(* IEC 61131-3 sources: STAR-PLC-Agent/results/raw/codex_matrix_resume_20261114/codex_deepseek/SELF010/functional/attempt_0001, 1 file *)

(* ---- test_program.st ---- *)
PROGRAM PLC_PRG
VAR
 BenchStep : UDINT := 0;
 BenchCalls : UDINT := 0;
 BenchDone : BOOL := FALSE;
 BenchUut0 : FB_Task;
 BenchUut1 : FB_Task;
 BenchUut2 : FB_Task;
 BenchUut3 : FB_Task;
 BenchUut4 : FB_Task;
 BenchUut5 : FB_Task;
 BenchUut6 : FB_Task;
 BenchUut7 : FB_Task;
 TraceIn_Fault : ARRAY[0..49] OF BOOL;
 TraceIn_Ack : ARRAY[0..49] OF BOOL;
 TraceIn_Reset : ARRAY[0..49] OF BOOL;
 TraceOut_Alarm : ARRAY[0..49] OF BOOL;
 TraceOut_Acknowledged : ARRAY[0..49] OF BOOL;
 TraceOut_Horn : ARRAY[0..49] OF BOOL;
END_VAR

IF NOT BenchDone THEN
 CASE BenchStep OF
 0:
   BenchUut0.Fault := FALSE;
   BenchUut0.Ack := FALSE;
   BenchUut0.Reset := FALSE;
   TraceIn_Fault[0] := BenchUut0.Fault;
   TraceIn_Ack[0] := BenchUut0.Ack;
   TraceIn_Reset[0] := BenchUut0.Reset;
   BenchUut0();
   TraceOut_Alarm[0] := BenchUut0.Alarm;
   TraceOut_Acknowledged[0] := BenchUut0.Acknowledged;
   TraceOut_Horn[0] := BenchUut0.Horn;
   BenchCalls := BenchCalls + 1;
 1:
   BenchUut0.Fault := TRUE;
   BenchUut0.Ack := TRUE;
   BenchUut0.Reset := FALSE;
   TraceIn_Fault[1] := BenchUut0.Fault;
   TraceIn_Ack[1] := BenchUut0.Ack;
   TraceIn_Reset[1] := BenchUut0.Reset;
   BenchUut0();
   TraceOut_Alarm[1] := BenchUut0.Alarm;
   TraceOut_Acknowledged[1] := BenchUut0.Acknowledged;
   TraceOut_Horn[1] := BenchUut0.Horn;
   BenchCalls := BenchCalls + 1;
 2:
   BenchUut0.Fault := TRUE;
   BenchUut0.Ack := TRUE;
   BenchUut0.Reset := FALSE;
   TraceIn_Fault[2] := BenchUut0.Fault;
   TraceIn_Ack[2] := BenchUut0.Ack;
   TraceIn_Reset[2] := BenchUut0.Reset;
   BenchUut0();
   TraceOut_Alarm[2] := BenchUut0.Alarm;
   TraceOut_Acknowledged[2] := BenchUut0.Acknowledged;
   TraceOut_Horn[2] := BenchUut0.Horn;
   BenchCalls := BenchCalls + 1;
 3:
   BenchUut0.Fault := FALSE;
   BenchUut0.Ack := FALSE;
   BenchUut0.Reset := FALSE;
   TraceIn_Fault[3] := BenchUut0.Fault;
   TraceIn_Ack[3] := BenchUut0.Ack;
   TraceIn_Reset[3] := BenchUut0.Reset;
   BenchUut0();
   TraceOut_Alarm[3] := BenchUut0.Alarm;
   TraceOut_Acknowledged[3] := BenchUut0.Acknowledged;
   TraceOut_Horn[3] := BenchUut0.Horn;
   BenchCalls := BenchCalls + 1;
 4:
   BenchUut0.Fault := TRUE;
   BenchUut0.Ack := FALSE;
   BenchUut0.Reset := FALSE;
   TraceIn_Fault[4] := BenchUut0.Fault;
   TraceIn_Ack[4] := BenchUut0.Ack;
   TraceIn_Reset[4] := BenchUut0.Reset;
   BenchUut0();
   TraceOut_Alarm[4] := BenchUut0.Alarm;
   TraceOut_Acknowledged[4] := BenchUut0.Acknowledged;
   TraceOut_Horn[4] := BenchUut0.Horn;
   BenchCalls := BenchCalls + 1;
 5:
   BenchUut0.Fault := FALSE;
   BenchUut0.Ack := FALSE;
   BenchUut0.Reset := TRUE;
   TraceIn_Fault[5] := BenchUut0.Fault;
   TraceIn_Ack[5] := BenchUut0.Ack;
   TraceIn_Reset[5] := BenchUut0.Reset;
   BenchUut0();
   TraceOut_Alarm[5] := BenchUut0.Alarm;
   TraceOut_Acknowledged[5] := BenchUut0.Acknowledged;
   TraceOut_Horn[5] := BenchUut0.Horn;
   BenchCalls := BenchCalls + 1;
 6:
   BenchUut1.Fault := TRUE;
   BenchUut1.Ack := FALSE;
   BenchUut1.Reset := TRUE;
   TraceIn_Fault[6] := BenchUut1.Fault;
   TraceIn_Ack[6] := BenchUut1.Ack;
   TraceIn_Reset[6] := BenchUut1.Reset;
   BenchUut1();
   TraceOut_Alarm[6] := BenchUut1.Alarm;
   TraceOut_Acknowledged[6] := BenchUut1.Acknowledged;
   TraceOut_Horn[6] := BenchUut1.Horn;
   BenchCalls := BenchCalls + 1;
 7:
   BenchUut1.Fault := TRUE;
   BenchUut1.Ack := TRUE;
   BenchUut1.Reset := TRUE;
   TraceIn_Fault[7] := BenchUut1.Fault;
   TraceIn_Ack[7] := BenchUut1.Ack;
   TraceIn_Reset[7] := BenchUut1.Reset;
   BenchUut1();
   TraceOut_Alarm[7] := BenchUut1.Alarm;
   TraceOut_Acknowledged[7] := BenchUut1.Acknowledged;
   TraceOut_Horn[7] := BenchUut1.Horn;
   BenchCalls := BenchCalls + 1;
 8:
   BenchUut1.Fault := FALSE;
   BenchUut1.Ack := TRUE;
   BenchUut1.Reset := TRUE;
   TraceIn_Fault[8] := BenchUut1.Fault;
   TraceIn_Ack[8] := BenchUut1.Ack;
   TraceIn_Reset[8] := BenchUut1.Reset;
   BenchUut1();
   TraceOut_Alarm[8] := BenchUut1.Alarm;
   TraceOut_Acknowledged[8] := BenchUut1.Acknowledged;
   TraceOut_Horn[8] := BenchUut1.Horn;
   BenchCalls := BenchCalls + 1;
 9:
   BenchUut2.Fault := TRUE;
   BenchUut2.Ack := FALSE;
   BenchUut2.Reset := TRUE;
   TraceIn_Fault[9] := BenchUut2.Fault;
   TraceIn_Ack[9] := BenchUut2.Ack;
   TraceIn_Reset[9] := BenchUut2.Reset;
   BenchUut2();
   TraceOut_Alarm[9] := BenchUut2.Alarm;
   TraceOut_Acknowledged[9] := BenchUut2.Acknowledged;
   TraceOut_Horn[9] := BenchUut2.Horn;
   BenchCalls := BenchCalls + 1;
 10:
   BenchUut2.Fault := TRUE;
   BenchUut2.Ack := TRUE;
   BenchUut2.Reset := TRUE;
   TraceIn_Fault[10] := BenchUut2.Fault;
   TraceIn_Ack[10] := BenchUut2.Ack;
   TraceIn_Reset[10] := BenchUut2.Reset;
   BenchUut2();
   TraceOut_Alarm[10] := BenchUut2.Alarm;
   TraceOut_Acknowledged[10] := BenchUut2.Acknowledged;
   TraceOut_Horn[10] := BenchUut2.Horn;
   BenchCalls := BenchCalls + 1;
 11:
   BenchUut2.Fault := TRUE;
   BenchUut2.Ack := TRUE;
   BenchUut2.Reset := TRUE;
   TraceIn_Fault[11] := BenchUut2.Fault;
   TraceIn_Ack[11] := BenchUut2.Ack;
   TraceIn_Reset[11] := BenchUut2.Reset;
   BenchUut2();
   TraceOut_Alarm[11] := BenchUut2.Alarm;
   TraceOut_Acknowledged[11] := BenchUut2.Acknowledged;
   TraceOut_Horn[11] := BenchUut2.Horn;
   BenchCalls := BenchCalls + 1;
 12:
   BenchUut3.Fault := FALSE;
   BenchUut3.Ack := TRUE;
   BenchUut3.Reset := FALSE;
   TraceIn_Fault[12] := BenchUut3.Fault;
   TraceIn_Ack[12] := BenchUut3.Ack;
   TraceIn_Reset[12] := BenchUut3.Reset;
   BenchUut3();
   TraceOut_Alarm[12] := BenchUut3.Alarm;
   TraceOut_Acknowledged[12] := BenchUut3.Acknowledged;
   TraceOut_Horn[12] := BenchUut3.Horn;
   BenchCalls := BenchCalls + 1;
 13:
   BenchUut3.Fault := TRUE;
   BenchUut3.Ack := FALSE;
   BenchUut3.Reset := FALSE;
   TraceIn_Fault[13] := BenchUut3.Fault;
   TraceIn_Ack[13] := BenchUut3.Ack;
   TraceIn_Reset[13] := BenchUut3.Reset;
   BenchUut3();
   TraceOut_Alarm[13] := BenchUut3.Alarm;
   TraceOut_Acknowledged[13] := BenchUut3.Acknowledged;
   TraceOut_Horn[13] := BenchUut3.Horn;
   BenchCalls := BenchCalls + 1;
 14:
   BenchUut3.Fault := FALSE;
   BenchUut3.Ack := FALSE;
   BenchUut3.Reset := FALSE;
   TraceIn_Fault[14] := BenchUut3.Fault;
   TraceIn_Ack[14] := BenchUut3.Ack;
   TraceIn_Reset[14] := BenchUut3.Reset;
   BenchUut3();
   TraceOut_Alarm[14] := BenchUut3.Alarm;
   TraceOut_Acknowledged[14] := BenchUut3.Acknowledged;
   TraceOut_Horn[14] := BenchUut3.Horn;
   BenchCalls := BenchCalls + 1;
 15:
   BenchUut3.Fault := FALSE;
   BenchUut3.Ack := TRUE;
   BenchUut3.Reset := FALSE;
   TraceIn_Fault[15] := BenchUut3.Fault;
   TraceIn_Ack[15] := BenchUut3.Ack;
   TraceIn_Reset[15] := BenchUut3.Reset;
   BenchUut3();
   TraceOut_Alarm[15] := BenchUut3.Alarm;
   TraceOut_Acknowledged[15] := BenchUut3.Acknowledged;
   TraceOut_Horn[15] := BenchUut3.Horn;
   BenchCalls := BenchCalls + 1;
 16:
   BenchUut3.Fault := TRUE;
   BenchUut3.Ack := TRUE;
   BenchUut3.Reset := FALSE;
   TraceIn_Fault[16] := BenchUut3.Fault;
   TraceIn_Ack[16] := BenchUut3.Ack;
   TraceIn_Reset[16] := BenchUut3.Reset;
   BenchUut3();
   TraceOut_Alarm[16] := BenchUut3.Alarm;
   TraceOut_Acknowledged[16] := BenchUut3.Acknowledged;
   TraceOut_Horn[16] := BenchUut3.Horn;
   BenchCalls := BenchCalls + 1;
 17:
   BenchUut3.Fault := TRUE;
   BenchUut3.Ack := FALSE;
   BenchUut3.Reset := TRUE;
   TraceIn_Fault[17] := BenchUut3.Fault;
   TraceIn_Ack[17] := BenchUut3.Ack;
   TraceIn_Reset[17] := BenchUut3.Reset;
   BenchUut3();
   TraceOut_Alarm[17] := BenchUut3.Alarm;
   TraceOut_Acknowledged[17] := BenchUut3.Acknowledged;
   TraceOut_Horn[17] := BenchUut3.Horn;
   BenchCalls := BenchCalls + 1;
 18:
   BenchUut3.Fault := FALSE;
   BenchUut3.Ack := FALSE;
   BenchUut3.Reset := TRUE;
   TraceIn_Fault[18] := BenchUut3.Fault;
   TraceIn_Ack[18] := BenchUut3.Ack;
   TraceIn_Reset[18] := BenchUut3.Reset;
   BenchUut3();
   TraceOut_Alarm[18] := BenchUut3.Alarm;
   TraceOut_Acknowledged[18] := BenchUut3.Acknowledged;
   TraceOut_Horn[18] := BenchUut3.Horn;
   BenchCalls := BenchCalls + 1;
 19:
   BenchUut4.Fault := TRUE;
   BenchUut4.Ack := FALSE;
   BenchUut4.Reset := FALSE;
   TraceIn_Fault[19] := BenchUut4.Fault;
   TraceIn_Ack[19] := BenchUut4.Ack;
   TraceIn_Reset[19] := BenchUut4.Reset;
   BenchUut4();
   TraceOut_Alarm[19] := BenchUut4.Alarm;
   TraceOut_Acknowledged[19] := BenchUut4.Acknowledged;
   TraceOut_Horn[19] := BenchUut4.Horn;
   BenchCalls := BenchCalls + 1;
 20:
   BenchUut4.Fault := FALSE;
   BenchUut4.Ack := FALSE;
   BenchUut4.Reset := FALSE;
   TraceIn_Fault[20] := BenchUut4.Fault;
   TraceIn_Ack[20] := BenchUut4.Ack;
   TraceIn_Reset[20] := BenchUut4.Reset;
   BenchUut4();
   TraceOut_Alarm[20] := BenchUut4.Alarm;
   TraceOut_Acknowledged[20] := BenchUut4.Acknowledged;
   TraceOut_Horn[20] := BenchUut4.Horn;
   BenchCalls := BenchCalls + 1;
 21:
   BenchUut4.Fault := FALSE;
   BenchUut4.Ack := TRUE;
   BenchUut4.Reset := FALSE;
   TraceIn_Fault[21] := BenchUut4.Fault;
   TraceIn_Ack[21] := BenchUut4.Ack;
   TraceIn_Reset[21] := BenchUut4.Reset;
   BenchUut4();
   TraceOut_Alarm[21] := BenchUut4.Alarm;
   TraceOut_Acknowledged[21] := BenchUut4.Acknowledged;
   TraceOut_Horn[21] := BenchUut4.Horn;
   BenchCalls := BenchCalls + 1;
 22:
   BenchUut4.Fault := FALSE;
   BenchUut4.Ack := FALSE;
   BenchUut4.Reset := FALSE;
   TraceIn_Fault[22] := BenchUut4.Fault;
   TraceIn_Ack[22] := BenchUut4.Ack;
   TraceIn_Reset[22] := BenchUut4.Reset;
   BenchUut4();
   TraceOut_Alarm[22] := BenchUut4.Alarm;
   TraceOut_Acknowledged[22] := BenchUut4.Acknowledged;
   TraceOut_Horn[22] := BenchUut4.Horn;
   BenchCalls := BenchCalls + 1;
 23:
   BenchUut4.Fault := FALSE;
   BenchUut4.Ack := FALSE;
   BenchUut4.Reset := TRUE;
   TraceIn_Fault[23] := BenchUut4.Fault;
   TraceIn_Ack[23] := BenchUut4.Ack;
   TraceIn_Reset[23] := BenchUut4.Reset;
   BenchUut4();
   TraceOut_Alarm[23] := BenchUut4.Alarm;
   TraceOut_Acknowledged[23] := BenchUut4.Acknowledged;
   TraceOut_Horn[23] := BenchUut4.Horn;
   BenchCalls := BenchCalls + 1;
 24:
   BenchUut4.Fault := FALSE;
   BenchUut4.Ack := FALSE;
   BenchUut4.Reset := FALSE;
   TraceIn_Fault[24] := BenchUut4.Fault;
   TraceIn_Ack[24] := BenchUut4.Ack;
   TraceIn_Reset[24] := BenchUut4.Reset;
   BenchUut4();
   TraceOut_Alarm[24] := BenchUut4.Alarm;
   TraceOut_Acknowledged[24] := BenchUut4.Acknowledged;
   TraceOut_Horn[24] := BenchUut4.Horn;
   BenchCalls := BenchCalls + 1;
 25:
   BenchUut4.Fault := FALSE;
   BenchUut4.Ack := TRUE;
   BenchUut4.Reset := FALSE;
   TraceIn_Fault[25] := BenchUut4.Fault;
   TraceIn_Ack[25] := BenchUut4.Ack;
   TraceIn_Reset[25] := BenchUut4.Reset;
   BenchUut4();
   TraceOut_Alarm[25] := BenchUut4.Alarm;
   TraceOut_Acknowledged[25] := BenchUut4.Acknowledged;
   TraceOut_Horn[25] := BenchUut4.Horn;
   BenchCalls := BenchCalls + 1;
 26:
   BenchUut5.Fault := FALSE;
   BenchUut5.Ack := FALSE;
   BenchUut5.Reset := FALSE;
   TraceIn_Fault[26] := BenchUut5.Fault;
   TraceIn_Ack[26] := BenchUut5.Ack;
   TraceIn_Reset[26] := BenchUut5.Reset;
   BenchUut5();
   TraceOut_Alarm[26] := BenchUut5.Alarm;
   TraceOut_Acknowledged[26] := BenchUut5.Acknowledged;
   TraceOut_Horn[26] := BenchUut5.Horn;
   BenchCalls := BenchCalls + 1;
 27:
   BenchUut5.Fault := TRUE;
   BenchUut5.Ack := TRUE;
   BenchUut5.Reset := FALSE;
   TraceIn_Fault[27] := BenchUut5.Fault;
   TraceIn_Ack[27] := BenchUut5.Ack;
   TraceIn_Reset[27] := BenchUut5.Reset;
   BenchUut5();
   TraceOut_Alarm[27] := BenchUut5.Alarm;
   TraceOut_Acknowledged[27] := BenchUut5.Acknowledged;
   TraceOut_Horn[27] := BenchUut5.Horn;
   BenchCalls := BenchCalls + 1;
 28:
   BenchUut5.Fault := TRUE;
   BenchUut5.Ack := TRUE;
   BenchUut5.Reset := FALSE;
   TraceIn_Fault[28] := BenchUut5.Fault;
   TraceIn_Ack[28] := BenchUut5.Ack;
   TraceIn_Reset[28] := BenchUut5.Reset;
   BenchUut5();
   TraceOut_Alarm[28] := BenchUut5.Alarm;
   TraceOut_Acknowledged[28] := BenchUut5.Acknowledged;
   TraceOut_Horn[28] := BenchUut5.Horn;
   BenchCalls := BenchCalls + 1;
 29:
   BenchUut5.Fault := FALSE;
   BenchUut5.Ack := FALSE;
   BenchUut5.Reset := FALSE;
   TraceIn_Fault[29] := BenchUut5.Fault;
   TraceIn_Ack[29] := BenchUut5.Ack;
   TraceIn_Reset[29] := BenchUut5.Reset;
   BenchUut5();
   TraceOut_Alarm[29] := BenchUut5.Alarm;
   TraceOut_Acknowledged[29] := BenchUut5.Acknowledged;
   TraceOut_Horn[29] := BenchUut5.Horn;
   BenchCalls := BenchCalls + 1;
 30:
   BenchUut5.Fault := TRUE;
   BenchUut5.Ack := FALSE;
   BenchUut5.Reset := FALSE;
   TraceIn_Fault[30] := BenchUut5.Fault;
   TraceIn_Ack[30] := BenchUut5.Ack;
   TraceIn_Reset[30] := BenchUut5.Reset;
   BenchUut5();
   TraceOut_Alarm[30] := BenchUut5.Alarm;
   TraceOut_Acknowledged[30] := BenchUut5.Acknowledged;
   TraceOut_Horn[30] := BenchUut5.Horn;
   BenchCalls := BenchCalls + 1;
 31:
   BenchUut5.Fault := FALSE;
   BenchUut5.Ack := FALSE;
   BenchUut5.Reset := TRUE;
   TraceIn_Fault[31] := BenchUut5.Fault;
   TraceIn_Ack[31] := BenchUut5.Ack;
   TraceIn_Reset[31] := BenchUut5.Reset;
   BenchUut5();
   TraceOut_Alarm[31] := BenchUut5.Alarm;
   TraceOut_Acknowledged[31] := BenchUut5.Acknowledged;
   TraceOut_Horn[31] := BenchUut5.Horn;
   BenchCalls := BenchCalls + 1;
 32:
   BenchUut5.Fault := TRUE;
   BenchUut5.Ack := FALSE;
   BenchUut5.Reset := TRUE;
   TraceIn_Fault[32] := BenchUut5.Fault;
   TraceIn_Ack[32] := BenchUut5.Ack;
   TraceIn_Reset[32] := BenchUut5.Reset;
   BenchUut5();
   TraceOut_Alarm[32] := BenchUut5.Alarm;
   TraceOut_Acknowledged[32] := BenchUut5.Acknowledged;
   TraceOut_Horn[32] := BenchUut5.Horn;
   BenchCalls := BenchCalls + 1;
 33:
   BenchUut5.Fault := TRUE;
   BenchUut5.Ack := FALSE;
   BenchUut5.Reset := TRUE;
   TraceIn_Fault[33] := BenchUut5.Fault;
   TraceIn_Ack[33] := BenchUut5.Ack;
   TraceIn_Reset[33] := BenchUut5.Reset;
   BenchUut5();
   TraceOut_Alarm[33] := BenchUut5.Alarm;
   TraceOut_Acknowledged[33] := BenchUut5.Acknowledged;
   TraceOut_Horn[33] := BenchUut5.Horn;
   BenchCalls := BenchCalls + 1;
 34:
   BenchUut6.Fault := FALSE;
   BenchUut6.Ack := FALSE;
   BenchUut6.Reset := FALSE;
   TraceIn_Fault[34] := BenchUut6.Fault;
   TraceIn_Ack[34] := BenchUut6.Ack;
   TraceIn_Reset[34] := BenchUut6.Reset;
   BenchUut6();
   TraceOut_Alarm[34] := BenchUut6.Alarm;
   TraceOut_Acknowledged[34] := BenchUut6.Acknowledged;
   TraceOut_Horn[34] := BenchUut6.Horn;
   BenchCalls := BenchCalls + 1;
 35:
   BenchUut6.Fault := TRUE;
   BenchUut6.Ack := TRUE;
   BenchUut6.Reset := FALSE;
   TraceIn_Fault[35] := BenchUut6.Fault;
   TraceIn_Ack[35] := BenchUut6.Ack;
   TraceIn_Reset[35] := BenchUut6.Reset;
   BenchUut6();
   TraceOut_Alarm[35] := BenchUut6.Alarm;
   TraceOut_Acknowledged[35] := BenchUut6.Acknowledged;
   TraceOut_Horn[35] := BenchUut6.Horn;
   BenchCalls := BenchCalls + 1;
 36:
   BenchUut6.Fault := TRUE;
   BenchUut6.Ack := TRUE;
   BenchUut6.Reset := FALSE;
   TraceIn_Fault[36] := BenchUut6.Fault;
   TraceIn_Ack[36] := BenchUut6.Ack;
   TraceIn_Reset[36] := BenchUut6.Reset;
   BenchUut6();
   TraceOut_Alarm[36] := BenchUut6.Alarm;
   TraceOut_Acknowledged[36] := BenchUut6.Acknowledged;
   TraceOut_Horn[36] := BenchUut6.Horn;
   BenchCalls := BenchCalls + 1;
 37:
   BenchUut6.Fault := FALSE;
   BenchUut6.Ack := FALSE;
   BenchUut6.Reset := FALSE;
   TraceIn_Fault[37] := BenchUut6.Fault;
   TraceIn_Ack[37] := BenchUut6.Ack;
   TraceIn_Reset[37] := BenchUut6.Reset;
   BenchUut6();
   TraceOut_Alarm[37] := BenchUut6.Alarm;
   TraceOut_Acknowledged[37] := BenchUut6.Acknowledged;
   TraceOut_Horn[37] := BenchUut6.Horn;
   BenchCalls := BenchCalls + 1;
 38:
   BenchUut6.Fault := TRUE;
   BenchUut6.Ack := FALSE;
   BenchUut6.Reset := FALSE;
   TraceIn_Fault[38] := BenchUut6.Fault;
   TraceIn_Ack[38] := BenchUut6.Ack;
   TraceIn_Reset[38] := BenchUut6.Reset;
   BenchUut6();
   TraceOut_Alarm[38] := BenchUut6.Alarm;
   TraceOut_Acknowledged[38] := BenchUut6.Acknowledged;
   TraceOut_Horn[38] := BenchUut6.Horn;
   BenchCalls := BenchCalls + 1;
 39:
   BenchUut6.Fault := FALSE;
   BenchUut6.Ack := FALSE;
   BenchUut6.Reset := TRUE;
   TraceIn_Fault[39] := BenchUut6.Fault;
   TraceIn_Ack[39] := BenchUut6.Ack;
   TraceIn_Reset[39] := BenchUut6.Reset;
   BenchUut6();
   TraceOut_Alarm[39] := BenchUut6.Alarm;
   TraceOut_Acknowledged[39] := BenchUut6.Acknowledged;
   TraceOut_Horn[39] := BenchUut6.Horn;
   BenchCalls := BenchCalls + 1;
 40:
   BenchUut6.Fault := FALSE;
   BenchUut6.Ack := TRUE;
   BenchUut6.Reset := TRUE;
   TraceIn_Fault[40] := BenchUut6.Fault;
   TraceIn_Ack[40] := BenchUut6.Ack;
   TraceIn_Reset[40] := BenchUut6.Reset;
   BenchUut6();
   TraceOut_Alarm[40] := BenchUut6.Alarm;
   TraceOut_Acknowledged[40] := BenchUut6.Acknowledged;
   TraceOut_Horn[40] := BenchUut6.Horn;
   BenchCalls := BenchCalls + 1;
 41:
   BenchUut6.Fault := FALSE;
   BenchUut6.Ack := TRUE;
   BenchUut6.Reset := TRUE;
   TraceIn_Fault[41] := BenchUut6.Fault;
   TraceIn_Ack[41] := BenchUut6.Ack;
   TraceIn_Reset[41] := BenchUut6.Reset;
   BenchUut6();
   TraceOut_Alarm[41] := BenchUut6.Alarm;
   TraceOut_Acknowledged[41] := BenchUut6.Acknowledged;
   TraceOut_Horn[41] := BenchUut6.Horn;
   BenchCalls := BenchCalls + 1;
 42:
   BenchUut7.Fault := FALSE;
   BenchUut7.Ack := FALSE;
   BenchUut7.Reset := FALSE;
   TraceIn_Fault[42] := BenchUut7.Fault;
   TraceIn_Ack[42] := BenchUut7.Ack;
   TraceIn_Reset[42] := BenchUut7.Reset;
   BenchUut7();
   TraceOut_Alarm[42] := BenchUut7.Alarm;
   TraceOut_Acknowledged[42] := BenchUut7.Acknowledged;
   TraceOut_Horn[42] := BenchUut7.Horn;
   BenchCalls := BenchCalls + 1;
 43:
   BenchUut7.Fault := TRUE;
   BenchUut7.Ack := TRUE;
   BenchUut7.Reset := FALSE;
   TraceIn_Fault[43] := BenchUut7.Fault;
   TraceIn_Ack[43] := BenchUut7.Ack;
   TraceIn_Reset[43] := BenchUut7.Reset;
   BenchUut7();
   TraceOut_Alarm[43] := BenchUut7.Alarm;
   TraceOut_Acknowledged[43] := BenchUut7.Acknowledged;
   TraceOut_Horn[43] := BenchUut7.Horn;
   BenchCalls := BenchCalls + 1;
 44:
   BenchUut7.Fault := TRUE;
   BenchUut7.Ack := TRUE;
   BenchUut7.Reset := FALSE;
   TraceIn_Fault[44] := BenchUut7.Fault;
   TraceIn_Ack[44] := BenchUut7.Ack;
   TraceIn_Reset[44] := BenchUut7.Reset;
   BenchUut7();
   TraceOut_Alarm[44] := BenchUut7.Alarm;
   TraceOut_Acknowledged[44] := BenchUut7.Acknowledged;
   TraceOut_Horn[44] := BenchUut7.Horn;
   BenchCalls := BenchCalls + 1;
 45:
   BenchUut7.Fault := FALSE;
   BenchUut7.Ack := FALSE;
   BenchUut7.Reset := FALSE;
   TraceIn_Fault[45] := BenchUut7.Fault;
   TraceIn_Ack[45] := BenchUut7.Ack;
   TraceIn_Reset[45] := BenchUut7.Reset;
   BenchUut7();
   TraceOut_Alarm[45] := BenchUut7.Alarm;
   TraceOut_Acknowledged[45] := BenchUut7.Acknowledged;
   TraceOut_Horn[45] := BenchUut7.Horn;
   BenchCalls := BenchCalls + 1;
 46:
   BenchUut7.Fault := TRUE;
   BenchUut7.Ack := FALSE;
   BenchUut7.Reset := FALSE;
   TraceIn_Fault[46] := BenchUut7.Fault;
   TraceIn_Ack[46] := BenchUut7.Ack;
   TraceIn_Reset[46] := BenchUut7.Reset;
   BenchUut7();
   TraceOut_Alarm[46] := BenchUut7.Alarm;
   TraceOut_Acknowledged[46] := BenchUut7.Acknowledged;
   TraceOut_Horn[46] := BenchUut7.Horn;
   BenchCalls := BenchCalls + 1;
 47:
   BenchUut7.Fault := FALSE;
   BenchUut7.Ack := FALSE;
   BenchUut7.Reset := TRUE;
   TraceIn_Fault[47] := BenchUut7.Fault;
   TraceIn_Ack[47] := BenchUut7.Ack;
   TraceIn_Reset[47] := BenchUut7.Reset;
   BenchUut7();
   TraceOut_Alarm[47] := BenchUut7.Alarm;
   TraceOut_Acknowledged[47] := BenchUut7.Acknowledged;
   TraceOut_Horn[47] := BenchUut7.Horn;
   BenchCalls := BenchCalls + 1;
 48:
   BenchUut7.Fault := FALSE;
   BenchUut7.Ack := FALSE;
   BenchUut7.Reset := FALSE;
   TraceIn_Fault[48] := BenchUut7.Fault;
   TraceIn_Ack[48] := BenchUut7.Ack;
   TraceIn_Reset[48] := BenchUut7.Reset;
   BenchUut7();
   TraceOut_Alarm[48] := BenchUut7.Alarm;
   TraceOut_Acknowledged[48] := BenchUut7.Acknowledged;
   TraceOut_Horn[48] := BenchUut7.Horn;
   BenchCalls := BenchCalls + 1;
 49:
   BenchUut7.Fault := FALSE;
   BenchUut7.Ack := FALSE;
   BenchUut7.Reset := FALSE;
   TraceIn_Fault[49] := BenchUut7.Fault;
   TraceIn_Ack[49] := BenchUut7.Ack;
   TraceIn_Reset[49] := BenchUut7.Reset;
   BenchUut7();
   TraceOut_Alarm[49] := BenchUut7.Alarm;
   TraceOut_Acknowledged[49] := BenchUut7.Acknowledged;
   TraceOut_Horn[49] := BenchUut7.Horn;
   BenchCalls := BenchCalls + 1;
 END_CASE;
 BenchStep := BenchStep + 1;
 IF BenchStep >= 50 THEN BenchDone := TRUE; END_IF;
END_IF;
END_PROGRAM
